Fanuc KAREL source: KD00052.KL

PROGRAM KD00052
%NOLOCKGROUP
%DEFGROUP = 1
VAR
  I: INTEGER
  J: INTEGER
  B: BOOLEAN
  R: REAL
  S: STRING[80]
  P: POSITION
BEGIN
  MOVE TO P,
  WHEN TIME 100 BEFORE NODE[1] DO DOUT[1] = TRUE
  ENDMOVE
END KD00052
